DATA_BLOCK "PressControl_DB"
{ S7_Optimized_Access := 'FALSE' }
VERSION : 0.1
NON_RETAIN
"PressControl"

BEGIN

END_DATA_BLOCK

